(*
SPDX-FileCopyrightText: © 2026 Oleksandr Tiutyk <trofimich@gmail.com>
SPDX-License-Identifier: MIT
License: https://opensource.org/license/mit
*)

(*!
<summary>Provides static helper methods for throwing FileSystem-specific exceptions.</summary>
<description>
Constructs stack-local template exceptions, formats diagnostics without heap allocation and propagates them
through ExceptionManager.
</description>
*)

PROGRAM FileSystemExceptions
VAR
	{attribute 'hide'} 
	_ClassName : STRING := __POUNAME();
END_VAR

//! <summary>Borrows the concrete class name for the lifetime of this instance; callers must not modify it.</summary>
{attribute 'monitoring' := 'call'}
PROPERTY ClassName : REFERENCE TO STRING
GET
ClassName REF= _ClassName;
END_GET
END_PROPERTY

//! <summary>Borrows the compiler-initialized namespace; callers must not modify the returned reference.</summary>
{attribute 'monitoring' := 'call'}
PROPERTY NamespaceName : REFERENCE TO STRING
GET
NamespaceName REF= CurrentNamespace.Name;
END_GET
END_PROPERTY

(*!
<summary>Raises a FileSystemException without requiring a caller-owned exception variable.</summary>
<description>Constructs a temporary stack template and delegates to FileSystemException.Throw.</description>
<param name="sourceNamespaceName">Namespace of the caller.</param>
<param name="sourceClassName">Class name of the caller.</param>
<param name="sourcePOUName">POU name of the caller.</param>
<param name="sourcePosition">Source position of the caller.</param>
<param name="message">Diagnostic explanation.</param>
<param name="errorCode">Native/ADS error code, or 0 if unassigned.</param>
*)
METHOD ThrowFileSystem
VAR_INPUT
	sourceNamespaceName : STRING;
	sourceClassName : STRING;
	sourcePOUName : STRING;
	sourcePosition : STRING;
END_VAR
VAR_IN_OUT CONSTANT
	message : TOF_Core.ERROR_MESSAGE;
END_VAR
VAR_INPUT
	errorCode : UDINT := 0;
END_VAR
VAR
	exception : FileSystemException;
END_VAR
exception.Throw(
	sourceNamespaceName := sourceNamespaceName,
	sourceClassName := sourceClassName,
	sourcePOUName := sourcePOUName,
	sourcePosition := sourcePosition,
	message := message,
	errorCode := errorCode
);
END_METHOD

(*!
<summary>Raises an InvalidPathException without requiring a caller-owned exception variable.</summary>
<description>Constructs a temporary stack template and delegates to InvalidPathException.Throw.</description>
<param name="sourceNamespaceName">Namespace of the caller.</param>
<param name="sourceClassName">Class name of the caller.</param>
<param name="sourcePOUName">POU name of the caller.</param>
<param name="sourcePosition">Source position of the caller.</param>
<param name="path">Rejected filesystem path.</param>
<param name="errorMessage">Diagnostic explanation.</param>
*)
METHOD ThrowInvalidPath
VAR_INPUT
	sourceNamespaceName : STRING;
	sourceClassName : STRING;
	sourcePOUName : STRING;
	sourcePosition : STRING;
END_VAR
VAR_IN_OUT CONSTANT
	path : STRING(255);
END_VAR
VAR_INPUT
	errorMessage : WSTRING(255);
END_VAR
VAR
	exception : InvalidPathException;
END_VAR
exception.Throw(
	sourceNamespaceName := sourceNamespaceName,
	sourceClassName := sourceClassName,
	sourcePOUName := sourcePOUName,
	sourcePosition := sourcePosition,
	path := path,
	errorMessage := errorMessage
);
END_METHOD

END_PROGRAM

(* stored: Version 1.1.0.1
   POU FileSystemExceptions: Id {dd62c6ab-3d90-4ca9-9192-7d723cc3b5f8}, SpecialFunc None
   Property ClassName: Id {9e8edd6f-741f-4c70-9a0e-92b145c6a8ce}
   Get Get: Id {cd6c45ad-5ba9-40f4-b5c9-1813fd79bc04}
   Property NamespaceName: Id {7e87426e-8aa4-4074-8621-d6b60cc67dbd}
   Get Get: Id {e2dcc754-d09d-452b-908a-f6078efd2def}
   Method ThrowFileSystem: Id {09d909ba-c131-4a7e-8485-2eace484a12d}
   Method ThrowInvalidPath: Id {cab3ac12-7ebf-48ed-a71e-7ca691e520c2} *)
